Fanuc KAREL source: KT00710.KL

PROGRAM KT00710
%NOLOCKGROUP
VAR
  B1: BOOLEAN
  B2: BOOLEAN
  OUT: BOOLEAN
BEGIN
  B1 = TRUE
  B2 = FALSE
  B1 = TRUE
  B2 = FALSE
  OUT = UNINIT(B1)
END KT00710
